{attribute 'qualified_only'}
{attribute 'strict'}
{attribute 'to_string'}
TYPE E_SafetyState :
(
	enum_RnD_2_Safe := 0,
	enum_Safe_2_RnD := 1,
	enum_RnD_2_Armed := 2,
	enum_Armed_2_RnD := 3
);
END_TYPE

(* stored: Version 1.1.0.1, ProductVersion 3.1.4026.18
   EnumerationTextList E_SafetyState: Id {7e58701e-5d58-4fc9-9499-789b690c2c97} *)
